Fanuc KAREL source: KA00124.KL

PROGRAM KA00124
%NOLOCKGROUP
VAR
  SRC: ARRAY[2] OF BYTE
  DST: STRING[80]
BEGIN
  SRC[1] = 2
  DST = SRC[1]
END KA00124
